(* IEC 61131-3 sources: Lasal-MCP/examples/SampleSource/LASALScreenAdvancedSolution/LASALScreenAdvancedSolution/LASALScreenAdvacnedSolution/Stations/MachineControl/MachineControl/Network/STDAlarm, 1 file *)

(* ---- ONE_STDAlarm_Table.st ---- *)
#define OBJECTS_CONFIG

#include "..\..\Class\_AlarmX0Para\_AlarmX0Para.h"
#include <.\lsl_st_mt.h>
#include "..\..\Class\_AlarmXBuffer\AlarmXBuffer.h"

FUNCTION GLOBAL TAB ONE_STDAlarm
-1$UINT, 0$UINT,
1$UINT, 0$UINT,

3$UDINT,
TO_UDINT(800276940), "_AlarmX0Para", 0$UINT, 11$UINT, 1$UINT,
TO_UDINT(2835625764), "_AlarmXBuffer", 0$UINT, 20$UINT, 1$UINT,
TO_UDINT(265160476), "UserAlarmGenerator", 1$UINT, 1$UINT, 1$UINT,

_NO_ATTR, TO_UDINT(3769593602), "BATTERIELOW_ERROR",

_NO_ATTR, TO_UDINT(3212185425), "_ALARMXBUFFER1",

_NO_ATTR, TO_UDINT(2488598847), "BATTERYALARM",

//Internal connections
0$UDINT,
0$UDINT,
0$UDINT,
1$UDINT,
TO_UDINT(2), "Out_alarm", TO_UDINT(0), "ClassSvr",

//Initialization values
0$UDINT,
4$UDINT,
TO_UDINT(0), "Config", TO_UDINT(0),//|STDAlarm.BatterieLow_Error.Config;
TO_UDINT(1), "No", TO_UDINT(500),//|STDAlarm._AlarmXBuffer1.No;
TO_UDINT(2), "In_status", TO_UDINT(0),//|STDAlarm.BatteryAlarm.In_status;
TO_UDINT(2), "In_mode", TO_UDINT(0),//|STDAlarm.BatteryAlarm.In_mode;

//Symbolic initialization values
0$UDINT,
0$UDINT,

//Initialization of string values
0$UDINT,
0$UDINT,

//Configuration of tasks (RealTime, Cyclic, Background)
0$UDINT,
0$UDINT,

0$UDINT,
1$UDINT,
TO_UDINT(2), (100)$UDINT, 4194303$DINT, 	//BATTERYALARM

0$UDINT,
0$UDINT,

//External connections
0$UDINT,
1$UDINT,
TO_UDINT(2), "In_status", C_DIR, TO_UDINT(3849002512), "STDPLC_InfoMC1","BatteryOk",

//Magic internal connections
0$UDINT,
0$UDINT,

//Configuration of timeslots of tasks (RealTime, Cyclic)
#ifdef __LSLLDR_TIMESLOTS__
0$UDINT,
0$UDINT,

0$UDINT,
0$UDINT,

#endif //__LSLLDR_TIMESLOTS__

//MultiMaster connections
#ifdef __LSLLDR_MULTIMASTER__
0$UDINT,
0$UDINT,
#endif //__LSLLDR_MULTIMASTER__

//Configuration for task ID (RealTime, CyclicTime)
#ifdef __LSLLDR_TASKID__
"\\\\TASKS2  "
0$UDINT,
0$UDINT,

0$UDINT,
1$UDINT,
(0)$UDINT, 	//BATTERYALARM

0$UDINT,
0$UDINT,

#endif //__LSLLDR_TASKID__

END_FUNCTION
